(* IEC 61131-3 sources: trust-platform/manual-tests/root-a/libs/Utils, 1 file *)

(* ---- Lib.st ---- *)
NAMESPACE Vendor.Utils
FUNCTION UtilFn : DINT
VAR_INPUT X : DINT; END_VAR
UtilFn := X;
END_FUNCTION
END_NAMESPACE
